TYPE coffee :
STRUCT

sName						: STRING;
fPrice						: REAL;
sIngredients				: STRING;


END_STRUCT
END_TYPE

(* stored: Version 1.1.0.1
   DUT coffee: Id {933616ed-3c5b-4965-8d7d-4b800fcc0dfc} *)
